Fanuc KAREL source: NC0001.KL

PROGRAM NC0001
%NOLOCKGROUP
ROUTINE R
VAR
  X : INTEGER
BEGIN
  X = 1
  X = X + 1
END R
BEGIN
  R
END NC0001
